// Mitsubishi GX Works2 project: 48_STRUCT_X1_Y1   PLC: FX3U/FX3UC

PROGRAM 1
(* structured ladder/FBD written out as ST: instructions are called as NAME(EN, inputs, outputs); _pN, _eN, _tN stand for wires *)
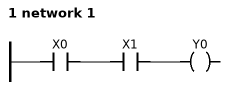
(* network 1 *)
Y0 := X0 AND X1;
END_PROGRAM
